// TIA Portal V20 export
DATA_BLOCK "Leuchtmelder Ampel_DB"   // DB77
// stored: InstanceOfName Leuchtmelder Ampel, InstanceOfType FB
"Leuchtmelder Ampel"
   // VAR
   //    Ampelbaustein_MG_Instance { S7_SetPoint := 'True'} : "Ampelbaustein_MG";
   //    OUT_Ampel_rot { S7_SetPoint := 'True'} : Bool;
   //    OUT_Ampel_gelb { S7_SetPoint := 'True'} : Bool;
   //    OUT_Ampel_gruen { S7_SetPoint := 'True'} : Bool;
   //    OUT_Akkustik { S7_SetPoint := 'True'} : Bool;
   // END_VAR
BEGIN
   Ampelbaustein_MG_Instance.Sammelstoerung := FALSE;
   Ampelbaustein_MG_Instance.BA_0 := FALSE;
   Ampelbaustein_MG_Instance.BA_A := FALSE;
   Ampelbaustein_MG_Instance.BA_M := TRUE;
   Ampelbaustein_MG_Instance.BA_R := FALSE;
   Ampelbaustein_MG_Instance.BA_V := FALSE;
   Ampelbaustein_MG_Instance.Ablauf_ist_aktiv := FALSE;
   Ampelbaustein_MG_Instance.Blinker := FALSE;
   Ampelbaustein_MG_Instance.Ampel_rot := FALSE;
   Ampelbaustein_MG_Instance.Ampel_gelb := FALSE;
   Ampelbaustein_MG_Instance.Ampel_gruen := FALSE;
   Ampelbaustein_MG_Instance.Akkustik := FALSE;
   Ampelbaustein_MG_Instance.Timer_Hupe_EIN.PT := T#5M;
   Ampelbaustein_MG_Instance.Timer_Hupe_EIN.IN := FALSE;
   Ampelbaustein_MG_Instance.Timer_Hupe_Aus.PT := T#10M;
   Ampelbaustein_MG_Instance.Timer_Hupe_Aus.IN := FALSE;
   Ampelbaustein_MG_Instance.Ampel_Zustand := 0;
END_DATA_BLOCK
